(* IEC 61131-3 sources: SortJet_MasterSPS_Aufbau.fbsproj/Device.device.xml.v3^/Plc Logic.plclogic.xml.v3^/Application.application.xml.v3^/09_Station/Stationen/Anlegetisch[201,205]/0_Konfig, 6 files *)

(* ---- Antriebsinformationen_201.gvl ---- *)
(* METADATA
{
	"v3Meta": {
		"objectGuid": "6db4b2f7-21ef-4267-9852-06546c6f86b1"
	}
}
*)
{attribute 'allow_unqualified_access'}
NAMESPACE Antriebsinformationen_201
VAR_GLOBAL

//-------------------------------------------------------------------------------------------------
// ANTRIEBSINFORMATION
//-------------------------------------------------------------------------------------------------

  apgInfoStation201Glastransport : ARRAY[cWAND_1..cANZAHL_WAENDE] OF AntriebsInformationen := [
    (
      wAchsID                                 :=     13,  // Achs ID aus dem EConSet
      stTyp                                   := 'Belt',  // Typ
      wpSchaltschrank                         :=   2010,  // Daten aus dem Schaltplan
      wpSchaltplanreihe                       :=      2,  // Daten aus dem Schaltplan
      wpSchaltplanseite                       :=    100,  // Daten aus dem Schaltplan
      rpMaxGeschwindigkeit                    :=   1000,  // [mm/s]   Max- Geschwindigkeit für den Automatikbetrieb
      rpHandGeschwindigkeit                   :=    200,  // [mm/s]   Hand- Geschwindigkeit
      rpReduzierteGeschwindigkeit             :=     67,  // [mm/s]   Reduzierte Geschwindigkeit
      rpReferenzGeschwindigkeit               :=      0,  // [mm/s]   Geschwindigkeit für die Referenzfahrt
      rpEinrichtGeschwindigkeit               :=     50,  // [mm/s]   Max Geschwindigkeit während der Einrichtung der Anlage
      rpMaxBeschleunigung                     :=   1500,  // [mm/s^2] Max Beschleunigung
      rpMaxVerzoegerung                       :=   2000,  // [mm/s^2] Max Verzoegerung
      rpMaxRuckzeit                           :=     50,  // [ms]     Ruckzeit des Antriebs
      rpReduzierteBeschleunigung              :=   1000,  // [mm/s^2] Reduzierte Beschleunigung
      rpReduzierteVerzoegerung                :=   1000,  // [mm/s^2] Reduzierte Verzoegerung
      rpBeschleunigungFremdanlage             :=   1000,  // [mm/s^2] Beschleunigung zu einer Fremdanlage
      rpGeschwindigkeitMessen                 :=    667,  // [mm/s] Geschwindigkeit beim Scheiben messen
      rpGeschwindigkeitSystemcheck            :=  500.0,  // [mm/s]   Geschwindigkeit im Systemcheck (nur Glastransport)
      rpGeschwindigkeitSystemcheckReduzierung :=  167.0,  // [mm/s]   Geschwindigkeit im Systemcheck bei belegtem Vorstop-Sensor (nur Glastransport)
      stOptionen                              := ( eEndschalterQuelle    := Endschalterquelle_EN.KEINE,     // Hardware-Endschalter: KEINE, UMRICHTER oder SPS
                                                   bVersorgungUeberXVR   := FALSE,                          // XVR-Modus: brueckt Hauptschalter 400 V und LS 230 V
                                                   bBremseLoesenFreigabe := FALSE )                         // Der Antrieb darf über eine Betriebsart die Bremse lösen
    )];

  apgInfoStation201Glastransport_Slave : ARRAY[cWAND_1..cANZAHL_WAENDE] OF AntriebsInformationen := [
    (
      wAchsID                                 :=     65,  // Achs ID aus dem EConSet
      stTyp                                   := 'BeltSl',  // Typ
      wpSchaltschrank                         :=      0,  // Daten aus dem Schaltplan
      wpSchaltplanreihe                       :=      2,  // Daten aus dem Schaltplan
      wpSchaltplanseite                       :=    100,  // Daten aus dem Schaltplan
      rpMaxGeschwindigkeit                    :=   1000,  // [mm/s]   Max- Geschwindigkeit für den Automatikbetrieb
      rpHandGeschwindigkeit                   :=    333,  // [mm/s]   Hand- Geschwindigkeit
      rpReduzierteGeschwindigkeit             :=    250,  // [mm/s]   Reduzierte Geschwindigkeit
      rpReferenzGeschwindigkeit               :=      0,  // [mm/s]   Geschwindigkeit für die Referenzfahrt
      rpEinrichtGeschwindigkeit               :=    100,  // [mm/s]   Max Geschwindigkeit während der Einrichtung der Anlage
      rpMaxBeschleunigung                     :=   1500,  // [mm/s^2] Max Beschleunigung
      rpMaxVerzoegerung                       :=   2000,  // [mm/s^2] Max Verzoegerung
      rpMaxRuckzeit                           :=     50,  // [ms]     Ruckzeit des Antriebs
      rpReduzierteBeschleunigung              :=    500,  // [mm/s^2] Reduzierte Beschleunigung
      rpReduzierteVerzoegerung                :=    500,  // [mm/s^2] Reduzierte Verzoegerung
      rpBeschleunigungFremdanlage             :=      0,  // [mm/s^2] Beschleunigung zu einer Fremdanlage
      rpGeschwindigkeitMessen                 :=   1000,  // [mm/s] Geschwindigkeit beim Scheiben messen
      rpGeschwindigkeitSystemcheck            :=  500.0,  // [mm/s]   Geschwindigkeit im Systemcheck (nur Glastransport)
      rpGeschwindigkeitSystemcheckReduzierung :=  167.0,  // [mm/s]   Geschwindigkeit im Systemcheck bei belegtem Vorstop-Sensor (nur Glastransport)
      stOptionen                              := ( eEndschalterQuelle    := Endschalterquelle_EN.KEINE,     // Hardware-Endschalter: KEINE, UMRICHTER oder SPS
                                                   bVersorgungUeberXVR   := FALSE,                          // XVR-Modus: brueckt Hauptschalter 400 V und LS 230 V
                                                   bBremseLoesenFreigabe := FALSE )                         // Der Antrieb darf über eine Betriebsart die Bremse lösen
    )];

  apgInfoStation201Messachse : AntriebsInformationen :=
    (
      wAchsID                                 :=        14,  // Achs ID aus dem EConSet
      stTyp                                   := 'Measure',  // Typ
      wpSchaltschrank                         :=      2011,  // Daten aus dem Schaltplan
      wpSchaltplanreihe                       :=         2,  // Daten aus dem Schaltplan
      wpSchaltplanseite                       :=       100,  // Daten aus dem Schaltplan
      rpMaxGeschwindigkeit                    :=      1000,  // [mm/s]   Max- Geschwindigkeit für den Automatikbetrieb
      rpHandGeschwindigkeit                   :=       333,  // [mm/s]   Hand- Geschwindigkeit
      rpReduzierteGeschwindigkeit             :=         0,  // [mm/s]   Reduzierte Geschwindigkeit
      rpReferenzGeschwindigkeit               :=        50,  // [mm/s]   Geschwindigkeit für die Referenzfahrt
      rpEinrichtGeschwindigkeit               :=         0,  // [mm/s]   Max Geschwindigkeit während der Einrichtung der Anlage
      rpMaxBeschleunigung                     :=      2500,  // [mm/s^2] Max Beschleunigung
      rpMaxVerzoegerung                       :=      2500,  // [mm/s^2] Max Verzoegerung
      rpMaxRuckzeit                           :=       500,  // [ms]     Ruckzeit des Antriebs
      rpReduzierteBeschleunigung              :=       500,  // [mm/s^2] Reduzierte Beschleunigung
      rpReduzierteVerzoegerung                :=       500,  // [mm/s^2] Reduzierte Verzoegerung
      rpBeschleunigungFremdanlage             :=         0,  // [mm/s^2] Beschleunigung zu einer Fremdanlage
      rpGeschwindigkeitMessen                 :=         0,  // [mm/s] Geschwindigkeit beim Scheiben messen
      rpGeschwindigkeitSystemcheck            :=     500.0,  // [mm/s]   Geschwindigkeit im Systemcheck (nur Glastransport)
      rpGeschwindigkeitSystemcheckReduzierung :=     167.0,  // [mm/s]   Geschwindigkeit im Systemcheck bei belegtem Vorstop-Sensor (nur Glastransport)
      stOptionen                              := ( eEndschalterQuelle    := Endschalterquelle_EN.UMRICHTER, // Hardware-Endschalter: KEINE, UMRICHTER oder SPS
                                                   bVersorgungUeberXVR   := FALSE,                          // XVR-Modus: brueckt Hauptschalter 400 V und LS 230 V
                                                   bBremseLoesenFreigabe := FALSE )                         // Der Antrieb darf über eine Betriebsart die Bremse lösen
    );

END_VAR

END_NAMESPACE

(* ---- Antriebsinformationen_205.gvl ---- *)
(* METADATA
{
	"v3Meta": {
		"objectGuid": "115b641a-a462-4b18-943b-f0d19b116a3d"
	}
}
*)
{attribute 'allow_unqualified_access'}
NAMESPACE Antriebsinformationen_205
VAR_GLOBAL

//-------------------------------------------------------------------------------------------------
// ANTRIEBSINFORMATION
//-------------------------------------------------------------------------------------------------

  apgInfoStation205Glastransport : ARRAY[cWAND_1..cANZAHL_WAENDE] OF AntriebsInformationen := [
    (
      wAchsID                                 :=     9,  // Achs ID aus dem EConSet
      stTyp                                   := 'Belt',  // Typ
      wpSchaltschrank                         :=   2050,  // Daten aus dem Schaltplan
      wpSchaltplanreihe                       :=      2,  // Daten aus dem Schaltplan
      wpSchaltplanseite                       :=    100,  // Daten aus dem Schaltplan
      rpMaxGeschwindigkeit                    :=   1000,  // [mm/s]   Max- Geschwindigkeit für den Automatikbetrieb
      rpHandGeschwindigkeit                   :=    200,  // [mm/s]   Hand- Geschwindigkeit
      rpReduzierteGeschwindigkeit             :=     67,  // [mm/s]   Reduzierte Geschwindigkeit
      rpReferenzGeschwindigkeit               :=      0,  // [mm/s]   Geschwindigkeit für die Referenzfahrt
      rpEinrichtGeschwindigkeit               :=     50,  // [mm/s]   Max Geschwindigkeit während der Einrichtung der Anlage
      rpMaxBeschleunigung                     :=   1500,  // [mm/s^2] Max Beschleunigung
      rpMaxVerzoegerung                       :=   2000,  // [mm/s^2] Max Verzoegerung
      rpMaxRuckzeit                           :=     50,  // [ms]     Ruckzeit des Antriebs
      rpReduzierteBeschleunigung              :=   1000,  // [mm/s^2] Reduzierte Beschleunigung
      rpReduzierteVerzoegerung                :=   1000,  // [mm/s^2] Reduzierte Verzoegerung
      rpBeschleunigungFremdanlage             :=   1000,  // [mm/s^2] Beschleunigung zu einer Fremdanlage
      rpGeschwindigkeitMessen                 :=    667,  // [mm/s] Geschwindigkeit beim Scheiben messen
      rpGeschwindigkeitSystemcheck            :=  500.0,  // [mm/s]   Geschwindigkeit im Systemcheck (nur Glastransport)
      rpGeschwindigkeitSystemcheckReduzierung :=  167.0,  // [mm/s]   Geschwindigkeit im Systemcheck bei belegtem Vorstop-Sensor (nur Glastransport)
      stOptionen                              := ( eEndschalterQuelle    := Endschalterquelle_EN.KEINE,     // Hardware-Endschalter: KEINE, UMRICHTER oder SPS
                                                   bVersorgungUeberXVR   := FALSE,                          // XVR-Modus: brueckt Hauptschalter 400 V und LS 230 V
                                                   bBremseLoesenFreigabe := FALSE )                         // Der Antrieb darf über eine Betriebsart die Bremse lösen
    )];

  apgInfoStation205Glastransport_Slave : ARRAY[cWAND_1..cANZAHL_WAENDE] OF AntriebsInformationen := [
    (
      wAchsID                                 :=     65,  // Achs ID aus dem EConSet
      stTyp                                   := 'BeltSl',  // Typ
      wpSchaltschrank                         :=      0,  // Daten aus dem Schaltplan
      wpSchaltplanreihe                       :=      2,  // Daten aus dem Schaltplan
      wpSchaltplanseite                       :=    100,  // Daten aus dem Schaltplan
      rpMaxGeschwindigkeit                    :=   1000,  // [mm/s]   Max- Geschwindigkeit für den Automatikbetrieb
      rpHandGeschwindigkeit                   :=    333,  // [mm/s]   Hand- Geschwindigkeit
      rpReduzierteGeschwindigkeit             :=    250,  // [mm/s]   Reduzierte Geschwindigkeit
      rpReferenzGeschwindigkeit               :=      0,  // [mm/s]   Geschwindigkeit für die Referenzfahrt
      rpEinrichtGeschwindigkeit               :=    100,  // [mm/s]   Max Geschwindigkeit während der Einrichtung der Anlage
      rpMaxBeschleunigung                     :=   1500,  // [mm/s^2] Max Beschleunigung
      rpMaxVerzoegerung                       :=   2000,  // [mm/s^2] Max Verzoegerung
      rpMaxRuckzeit                           :=     50,  // [ms]     Ruckzeit des Antriebs
      rpReduzierteBeschleunigung              :=    500,  // [mm/s^2] Reduzierte Beschleunigung
      rpReduzierteVerzoegerung                :=    500,  // [mm/s^2] Reduzierte Verzoegerung
      rpBeschleunigungFremdanlage             :=      0,  // [mm/s^2] Beschleunigung zu einer Fremdanlage
      rpGeschwindigkeitMessen                 :=   1000,  // [mm/s] Geschwindigkeit beim Scheiben messen
      rpGeschwindigkeitSystemcheck            :=  500.0,  // [mm/s]   Geschwindigkeit im Systemcheck (nur Glastransport)
      rpGeschwindigkeitSystemcheckReduzierung :=  167.0,  // [mm/s]   Geschwindigkeit im Systemcheck bei belegtem Vorstop-Sensor (nur Glastransport)
      stOptionen                              := ( eEndschalterQuelle    := Endschalterquelle_EN.KEINE,     // Hardware-Endschalter: KEINE, UMRICHTER oder SPS
                                                   bVersorgungUeberXVR   := FALSE,                          // XVR-Modus: brueckt Hauptschalter 400 V und LS 230 V
                                                   bBremseLoesenFreigabe := FALSE )                         // Der Antrieb darf über eine Betriebsart die Bremse lösen
    )];

  apgInfoStation205Messachse : AntriebsInformationen :=
    (
      wAchsID                                 :=        10,  // Achs ID aus dem EConSet
      stTyp                                   := 'Measure',  // Typ
      wpSchaltschrank                         :=      2051,  // Daten aus dem Schaltplan
      wpSchaltplanreihe                       :=         2,  // Daten aus dem Schaltplan
      wpSchaltplanseite                       :=       100,  // Daten aus dem Schaltplan
      rpMaxGeschwindigkeit                    :=      1000,  // [mm/s]   Max- Geschwindigkeit für den Automatikbetrieb
      rpHandGeschwindigkeit                   :=       333,  // [mm/s]   Hand- Geschwindigkeit
      rpReduzierteGeschwindigkeit             :=         0,  // [mm/s]   Reduzierte Geschwindigkeit
      rpReferenzGeschwindigkeit               :=        50,  // [mm/s]   Geschwindigkeit für die Referenzfahrt
      rpEinrichtGeschwindigkeit               :=         0,  // [mm/s]   Max Geschwindigkeit während der Einrichtung der Anlage
      rpMaxBeschleunigung                     :=      2500,  // [mm/s^2] Max Beschleunigung
      rpMaxVerzoegerung                       :=      2500,  // [mm/s^2] Max Verzoegerung
      rpMaxRuckzeit                           :=       500,  // [ms]     Ruckzeit des Antriebs
      rpReduzierteBeschleunigung              :=       500,  // [mm/s^2] Reduzierte Beschleunigung
      rpReduzierteVerzoegerung                :=       500,  // [mm/s^2] Reduzierte Verzoegerung
      rpBeschleunigungFremdanlage             :=         0,  // [mm/s^2] Beschleunigung zu einer Fremdanlage
      rpGeschwindigkeitMessen                 :=         0,  // [mm/s] Geschwindigkeit beim Scheiben messen
      rpGeschwindigkeitSystemcheck            :=     500.0,  // [mm/s]   Geschwindigkeit im Systemcheck (nur Glastransport)
      rpGeschwindigkeitSystemcheckReduzierung :=     167.0,  // [mm/s]   Geschwindigkeit im Systemcheck bei belegtem Vorstop-Sensor (nur Glastransport)
      stOptionen                              := ( eEndschalterQuelle    := Endschalterquelle_EN.UMRICHTER, // Hardware-Endschalter: KEINE, UMRICHTER oder SPS
                                                   bVersorgungUeberXVR   := FALSE,                          // XVR-Modus: brueckt Hauptschalter 400 V und LS 230 V
                                                   bBremseLoesenFreigabe := FALSE )                         // Der Antrieb darf über eine Betriebsart die Bremse lösen
    );

END_VAR

END_NAMESPACE

(* ---- MK_Station_201.gvl ---- *)
(* METADATA
{
	"v3Meta": {
		"objectGuid": "3c311fcf-86c3-480c-8d89-6d8c270ee569"
	}
}
*)
{attribute 'allow_unqualified_access'}
NAMESPACE MK_Station_201
VAR_GLOBAL

//-------------------------------------------------------------------------------------------------
// MASCHINEPARAMETER: ANLEGETISCH
//-------------------------------------------------------------------------------------------------

  apgMKStation201 : Parameter_Station :=
    (
      stStationsNummern                     := ( NummerIntern :=   201,                                                      // Stationsnummer fuer das MMI und die Stationsangabe der Meldungen
                                                 NummerExtern :=  1201,                                                      // Stationsnummer fuer Bedienermeldungen
                                                 NummerSPS    :=   201 ),                                                    // Stationsnummer SPS-intern (Indizes)
      bDeaktivieren                         := FALSE,                                                                        // Station deaktiviert (keine Auftraege, keine Referenzfahrt)
      wMeldungsNummer                       := 1700,                                                                         // Basis-Meldungsnummer (WatchIO)
      eStationsTyp                          := eStation,                                                                     // Typ der Station
      eaAutomatikkreis                      := [eAutomatikkreis_1],                                                          // Automatikkreise, zu denen die Station gehoert
      eaSicherheitskreis                    := [eSicherheitskreis_2],                                                        // Sicherheitskreise, in die die Station eingebunden ist
      // astSicherheitskreisTeilabschaltung
      eSystemcheckZyklus                    := eSystemcheckZyklus_1,                                                         // In welchem Zyklus des Systemchecks die Station geprueft wird
      stSchnittstellendaten                 := ( wVorgaengerStation := cSTATION_DEFAULT,                                     // Station vor dieser Station (cSTATION_DYNAMISCH bei mehreren)
                                                 wNachfolgerStation := cSTATION_202,                                         // Station nach dieser Station (cSTATION_DYNAMISCH bei mehreren)
                                                 bStationIstShuttle := FALSE                                                 // Station ist ein Shuttle
                                               ),
      stStationsOptionen                    := ( stSystemcheck   :=  ( bScheibenVermessenSystemCheck               := TRUE,  // Scheiben im Systemcheck vermessen
                                                                       bScheibeNachSystemcheckAufAuslauf           := FALSE, // Scheibe nach dem Systemcheck auf den Auslaufsensor fahren
                                                                       bSystemCheckMitVorgaengerBatchTransport     := FALSE, // derzeit ohne Funktion
                                                                       bSystemCheckMitNachfolgerBatchTransport     := FALSE, // derzeit ohne Funktion
                                                                       bOptionSystemCheckScheibeMittigLegen        := FALSE  // derzeit ohne Funktion
                                                                     ),
                                                 stAnlegetisch   :=  (
                                                                       bIstAnlegestation                         := TRUE,    // Station an der Scheiben angelegt werden [Anlegetisch, Anlegewand]; im Systemcheck-Verbund nur mit genau einer Scheibe
                                                                       bAnschlagAutomatischAusfahren             := TRUE,    // Anschlaege beim Anlegen automatisch ausfahren (Vorgabe, am Taster umschaltbar)
                                                                       bAnlegetischMitEintransportVorgaenger     := FALSE    // VSG: Station entscheidet selbst zwischen Eintransport vom Vorgaenger und Anlegen
                                                                     ),
                                                 // stTransfershuttle
                                                 stGlastransport :=  ( bVortransport                             := FALSE,   // Vortransport aktivieren [Bsp.: Nach einem Eintransport mit gesetztem Bit <Letzte Scheibe>]
                                                                       bTransportMasterSlaveEintransport         := FALSE,   // derzeit ohne Funktion
                                                                       bTransportMasterSlaveAustransport         := TRUE,    // Austransport als Slave auf die Achse des Nachfolgers
                                                                       bGLasUebernahmeSenkrecht                  := FALSE,   // RKT - Eintransport in Senkrechter-Position bzw. in Waagerechter- Position [default]
                                                                       bAustransportISOLinie                     := FALSE,   // Austransport an eine ISO-Linie
                                                                       bScheibenVermessen                        := TRUE,    // Scheibenmessung am Anlegetisch/Anlegewand
                                                                       bMessrichtungNegativ                      := FALSE,   // Negative Fahrtrichtung beim Messen
                                                                       bScheibenmessungEintransport              := FALSE,   // Scheibenmessung beim Eintransport
                                                                       bScheibenmessungSensorVorabAuslauf        := FALSE    // Scheibenmessung mit SensorVorabAuslauf z.B. Anlegewand
                                                                      ),
                                                 // stEckuebergabe
                                                 // stDrehstation
                                                 bVorAbKomponentenAnsteuerung              := FALSE,                         // VorAbKomponentenAnsteuerung Auftraege werden bearbeitet
                                                 bVerstellungEinAusGefahrenLogikDrehen     := FALSE,                         // Verstellung: Logik ein-/ausgefahren gedreht
                                                 bLangsamfahrtNockenQuerfahrtAktivieren    := FALSE,                         // Querfahrt: Langsamfahrt-Nocken auswerten
                                                 bSKBlockierenDurchVorabSensoren           := FALSE,                         // Vorab-Sensoren belegt blockieren das Oeffnen des Sicherheitskreises
                                                 bStationLeerfahrenBeiSkAnforderung        := FALSE,                         // Station bei Anforderung Sicherheitskreis leerfahren
                                                 bGlasAbgenommenAutomatischQuittieren      := FALSE,                         // derzeit ohne Funktion
                                                 bScheibeAbnehmenNachEintransport          := FALSE                          // Scheibe nach dem Eintransport wieder abnehmen
                                               ),
      stStationsAufbau                      := ( bGeblase                      := [ cANZAHL_WAENDE(TRUE) ],                  // Ausbaustufe: Geblaese je Wand
                                                 bGlastransport                := [ cANZAHL_WAENDE(TRUE) ],                  // Ausbaustufe: Glastransport je Wand
                                                 bKippen                       := [ cANZAHL_WAENDE(TRUE) ],                  // Ausbaustufe: Kippen je Wand (Kipptisch 201 laut E-Plan)
                                                 bKippenSchuetz                := FALSE,                                     // Kippen ueber Schuetz statt Umrichter
                                                 bTransportVerstellung         := [ cANZAHL_WAENDE(FALSE) ],                 // Ausbaustufe Shuttle: Transport-/Dickenverstellung je Wand
                                                 bHub                          := FALSE,                                     // Ausbaustufe: Hub der Station
                                                 bHubrahmen                    := TRUE,                                      // Ausbaustufe: Hubrahmen (Riemen heben/senken)
                                                 bDrehen                       := FALSE,                                     // Ausbaustufe: Drehen
                                                 bQuerachse                    := FALSE,                                     // Ausbaustufe: Querachse
                                                 bMessachse                    := TRUE,                                      // Ausbaustufe: Messachse (Anlegetisch, Anlegewand)
                                                 bDruckluft                    := TRUE,                                      // Druckluftueberwachung vorhanden
                                                 bAnschlag                     := TRUE,                                      // Ausbaustufe: Ausrichtanschlaege
                                                 bSensorAuslauf                := TRUE,                                      // Auslaufsensor vorhanden
                                                 bSensorEinlauf                := TRUE,                                      // Einlaufsensor vorhanden
                                                 bSensorEinlaufStopp           := FALSE,                                     // Shuttle: zusaetzlicher Stopp-Sensor am Einlauf (ohne: Einlaufsensor), Gegenstueck zum Auslauf-Stopp im Rueckwaertstransport
                                                 bSensorAuslaufStopp           := FALSE,                                     // Shuttle: zusaetzlicher Stopp-Sensor am Auslauf (ohne: Auslaufsensor), Verfahrfreigabe und Scheibe hat Shuttle verlassen
                                                 bDurchlaufSperreZumNachfolger := FALSE,                                     // Ausbaustufe: bewegliche Abschrankung zum Nachfolger
                                                 bQuerfahrt                    := FALSE,                                     // Ausbaustufe: Querfahrt
                                                 bKipparme                     := FALSE,                                     // Ausbaustufe: Kipparme
                                                 bSlaveAntrieb                 := FALSE,                                     // Glastransport mit Slave-Antrieb
                                                 bMessachseAmEndeVomTisch      := FALSE,                                     // Messachse am Ende des Tisches (Hoehenfehler fragt den Bediener)
                                                 bWandverstellung              := [ FALSE ],                                 // Ausbaustufe Station: Wandverstellung je Wand
                                                 bWandverstellungMotorisch     := FALSE,                                     // Shuttle: Transport-/Wandverstellung mit Antrieb statt pneumatisch
                                                 bRoellchenleiste              := [ FALSE ],                                 // Ausbaustufe Station: Roellchenleiste je Wand
                                                 bDurchgang                    := FALSE,                                     // Station ist Teil eines Durchgangs (belegt = Oeffnen blockiert)
                                                 bRolltor                      := FALSE,                                     // Ausbaustufe Faecherwagen: Rolltor
                                                 bKlemmzylinder                := FALSE,                                     // Ausbaustufe Faecherwagen: Klemmzylinder fixiert den Oberrahmen beim Ein- und Ausschleusen
                                                 bGreifer                      := [cANZAHL_WAENDE(FALSE)],                   // Shuttle: Greifer je Wand (Scheibe aus dem Faecherwagen ziehen bzw. hineinschieben)
                                                 bRFID                         := FALSE,                                     // RFID-Leser vorhanden
                                                 bAGV                          := FALSE,                                     // Ausbaustufe Faecherwagen: Betrieb mit AGV
                                                 bDLSSchmiersystem             := FALSE,                                     // Zentralschmierung DLS vorhanden
                                                 bGlastransportSlaveVorhanden  := FALSE,                                     // Glastransport mit Slave-Antrieb (Meldungen/Ueberwachung Slave)
                                                 wHydraulikstation             := 0                                          // Faecherwagen Hydraulik: zugeordnete Hydraulikstation (cHYDRAULIKSTATION_x), 0 = keine
                                               ),
      stStationsParameter                   := ( rLaengeUebergroesseScheibe              := 4240,                            // Shuttle: ab dieser Scheibenlaenge gilt die Scheibe als uebergross [mm]
                                                 rMinGlasHoeheAutomatischenEintransport  := 500,                             // VSG: Mindesthoehe fuer automatischen Eintransport [mm]
                                                 rMinGlasLaengeAutomatischenEintransport := 500,                             // VSG: Mindestlaenge fuer automatischen Eintransport [mm]
                                                 wMaximaleAnzahlAktiverAuftraege         := 1,                               // derzeit ohne Funktion
                                                 rMinPosSwEsEingrenzung                  := 0.0,                             // Externer zusaetzlicher Software-Endschalter MIN; 0 = inaktiv; darf den MK-MIN nur weiter eingrenzen
                                                 rMaxPosSwEsEingrenzung                  := 0.0,                             // Externer zusaetzlicher Software-Endschalter MAX; 0 = inaktiv; darf den MK-MAX nur weiter eingrenzen
                                                 rPosFreigabePufferAusfahren             := 0.0                              // derzeit ohne Funktion
                                              ),
      // stFremdanlage
      stGlasdaten                           := [(
                                                 rlMinGlasLaenge                  := 350,                                    // minimal zulässige GlasLänge
                                                 rlMaxGlasLaenge                  := 2500,                                   // maximale zulässige GlasLänge
                                                 rlMinGlasHoehe                   := 190,                                    // minimal zulässige GlasHöhe
                                                 rlMaxGlasHoehe                   := 1800,                                   // maximale zulässige GlasHöhe
                                                 rlMinGlasDicke                   := 3,                                    // minimal zulässige GlasDicke
                                                 rlMaxGlasDicke                   := 12.76,                                     // maximal zulaessige Glasdicke [mm]
                                                 rlLaengeMaxGlas                  := 0.0                                     // maximal zulaessige Glaslaenge [mm]
                                               )]
      // astShuttleAnhaltenQuellen
    );

  apgMKStation201Glastransport : ARRAY[cWAND_1..cANZAHL_WAENDE] OF Parameter_Glastransport := [
    (
      rLaengeStation                        := 3200, // Länge der Station
      rScheibenabstand                      :=  300, // Der Abstand zwischen zwei Scheiben auf der Station
      rWegUeberEinlauf                      :=   50, // Weg ueber den Einlaufsensor hinaus [mm]
      rWegUeberAuslauf                      :=   50, // Weg ueber den Auslaufsensor hinaus [mm]
      rWegUeberSensorenSystemCheck          :=   15, // Der Weg der Ueber ein die Sensoren zum vermessen der Scheiben
      rUeberwachungAuslaufsensor            :=  500, // Ueberwachung des Auslaufsensors [Strecke in der der Auslaufsensor Frei / ueberfahren werden soll]
      rUeberwachungEinlaufsensor            :=  500, // Ueberwachung des Einlaufsensors [Strecke in der der Einlaufsensor Frei / ueberfahren werden soll]
      rWegUeberEinlaufEintransport          :=  150, // Eintransport vorwaerts: Abstand Scheibenhinterkante zum Einlaufsensor [mm]
      rWegUeberEinlaufAustransport          :=   50, // Lage Auf Einlauf: Scheibe liegt um diesen Weg auf dem Einlaufsensor [mm]
      rWegUeberAuslaufEintransport          :=   50, // Eintransport rueckwaerts: Abstand Scheibenhinterkante zum Auslaufsensor [mm]
      rWegUeberAuslaufAustransport          :=   50, // Lage Auf Auslauf: Weg ueber den Auslaufsensor hinaus [mm]
      rWegEinlaufsensorZuVorStopSensor      := 3100, // Beschreibt den Weg vum eine Scheibe beim EIntransport vom Einlaufsensor bis ueberden Vorabstopsensor zu verfahren
      rMesstoleranz                         :=   10, // Toleranz-Mass fuer die Scheibenlaengenmessung
      rMessstrecke                          := 3140, // Beschreibt die Strecke ziwischen 2 Sensoren die der Antrieb verfaehrt
      rWegstreckeBisZurVerzoegerung         := 2600  // Beschreibt die Strecke die gefahren werden soll bis der Antrieb abgebremst werden soll, dies gilt fuer Eintransportauftraege die das Bit "Letzte Scheibe" gesetzt haben
    )];

  apgMKStation201Messachse : Parameter_Messachse :=
    (
      rPositionUeberScheibenhoehe           :=      0, // Position der Zentrierleiste ueber dem Glas so dass das Glas angelegt werden kann
      rKorrekturOffset                      :=      0, // Korrektur der Position um einen Bestimmten Wert (Offset)
      rStreckePositionieren                 :=      0, // ?
      rVerfahrbereichsOffset                :=      0, // Korrektur des Verfahrens wenn
      rOffsetMessung                        :=      0, // ?
      rToleranz                             :=     10, // Toleranzwert in der Ausmessung der Höhe
      rAbstandSensorenOberUndUnterkante     :=    153, // Rechnerischer Abstand zwischen dem Sensor der die Scheibenunterkante misst und dem Sensor der die Scheibenoberkante misst
      rKorrekturOffsetVSGEintransport       := 0.0,    // Korrektur der Position um einen Bestimmten Wert (Offset) beim Eintransport von VSG
      rOffsetNullLinie                      := 0.0     // Offset das auf den Wert des Abstands zur Null-Linie aufgerechnet wird, um dies evtl zu korrigieren
    );

END_VAR
END_NAMESPACE

(* ---- MK_Station_205.gvl ---- *)
(* METADATA
{
	"v3Meta": {
		"objectGuid": "7b970d81-93e6-42b4-b0eb-c486128876da"
	}
}
*)
{attribute 'allow_unqualified_access'}
NAMESPACE MK_Station_205
VAR_GLOBAL

//-------------------------------------------------------------------------------------------------
// MASCHINEPARAMETER: ANLEGETISCH
//-------------------------------------------------------------------------------------------------

  apgMKStation205 : Parameter_Station :=
    (
      stStationsNummern                     := ( NummerIntern :=   205,                                                      // Stationsnummer fuer das MMI und die Stationsangabe der Meldungen
                                                 NummerExtern :=  1205,                                                      // Stationsnummer fuer Bedienermeldungen
                                                 NummerSPS    :=   205 ),                                                    // Stationsnummer SPS-intern (Indizes)
      bDeaktivieren                         := FALSE,                                                                         // Station deaktiviert (keine Auftraege, keine Referenzfahrt)
      wMeldungsNummer                       := 1760,                                                                         // Basis-Meldungsnummer (WatchIO)
      eStationsTyp                          := eStation,                                                                     // Typ der Station
      eaAutomatikkreis                      := [eAutomatikkreis_1],                                                          // Automatikkreise, zu denen die Station gehoert
      eaSicherheitskreis                    := [eSicherheitskreis_Undefiniert],                                              // Sicherheitskreise, in die die Station eingebunden ist
      // astSicherheitskreisTeilabschaltung
      eSystemcheckZyklus                    := eSystemcheckZyklus_1,                                                         // In welchem Zyklus des Systemchecks die Station geprueft wird
      stSchnittstellendaten                 := ( wVorgaengerStation := cSTATION_501,                                         // Station vor dieser Station (cSTATION_DYNAMISCH bei mehreren)
                                                 wNachfolgerStation := cSTATION_204,                                         // Station nach dieser Station (cSTATION_DYNAMISCH bei mehreren)
                                                 bStationIstShuttle := FALSE                                                 // Station ist ein Shuttle
                                               ),
      stStationsOptionen                    := ( stSystemcheck   :=  ( bScheibenVermessenSystemCheck               := TRUE,  // Scheiben im Systemcheck vermessen
                                                                       bScheibeNachSystemcheckAufAuslauf           := FALSE, // Scheibe nach dem Systemcheck auf den Auslaufsensor fahren
                                                                       bSystemCheckMitVorgaengerBatchTransport     := FALSE, // derzeit ohne Funktion
                                                                       bSystemCheckMitNachfolgerBatchTransport     := FALSE, // derzeit ohne Funktion
                                                                       bOptionSystemCheckScheibeMittigLegen        := FALSE  // derzeit ohne Funktion
                                                                     ),
                                                 stAnlegetisch   :=  (
                                                                       bIstAnlegestation                         := TRUE,    // Station an der Scheiben angelegt werden [Anlegetisch, Anlegewand]; im Systemcheck-Verbund nur mit genau einer Scheibe
                                                                       bAnschlagAutomatischAusfahren             := TRUE,    // Anschlaege beim Anlegen automatisch ausfahren (Vorgabe, am Taster umschaltbar)
                                                                       bAnlegetischMitEintransportVorgaenger     := TRUE     // VSG: Station entscheidet selbst zwischen Eintransport vom Vorgaenger und Anlegen
                                                                     ),
                                                 // stTransfershuttle
                                                 stGlastransport :=  ( bVortransport                             := FALSE,   // Vortransport aktivieren [Bsp.: Nach einem Eintransport mit gesetztem Bit <Letzte Scheibe>]
                                                                       bTransportMasterSlaveEintransport         := FALSE,   // derzeit ohne Funktion
                                                                       bTransportMasterSlaveAustransport         := TRUE,    // Austransport als Slave auf die Achse des Nachfolgers
                                                                       bGLasUebernahmeSenkrecht                  := FALSE,   // RKT - Eintransport in Senkrechter-Position bzw. in Waagerechter- Position [default]
                                                                       bAustransportISOLinie                     := FALSE,   // Austransport an eine ISO-Linie
                                                                       bScheibenVermessen                        := TRUE,    // Scheibenmessung am Anlegetisch/Anlegewand
                                                                       bMessrichtungNegativ                      := FALSE,   // Negative Fahrtrichtung beim Messen
                                                                       bScheibenmessungEintransport              := FALSE,   // Scheibenmessung beim Eintransport
                                                                       bScheibenmessungSensorVorabAuslauf        := FALSE    // Scheibenmessung mit SensorVorabAuslauf z.B. Anlegewand
                                                                      ),
                                                 // stEckuebergabe
                                                 // stDrehstation
                                                 bVorAbKomponentenAnsteuerung              := FALSE,                         // VorAbKomponentenAnsteuerung Auftraege werden bearbeitet
                                                 bVerstellungEinAusGefahrenLogikDrehen     := FALSE,                         // Verstellung: Logik ein-/ausgefahren gedreht
                                                 bLangsamfahrtNockenQuerfahrtAktivieren    := FALSE,                         // Querfahrt: Langsamfahrt-Nocken auswerten
                                                 bSKBlockierenDurchVorabSensoren           := FALSE,                         // Vorab-Sensoren belegt blockieren das Oeffnen des Sicherheitskreises
                                                 bStationLeerfahrenBeiSkAnforderung        := FALSE,                         // Station bei Anforderung Sicherheitskreis leerfahren
                                                 bGlasAbgenommenAutomatischQuittieren      := FALSE,                         // derzeit ohne Funktion
                                                 bScheibeAbnehmenNachEintransport          := FALSE                          // Scheibe nach dem Eintransport wieder abnehmen
                                               ),
      stStationsAufbau                      := ( bGeblase                      := [ cANZAHL_WAENDE(TRUE) ],                  // Ausbaustufe: Geblaese je Wand
                                                 bGlastransport                := [ cANZAHL_WAENDE(TRUE) ],                  // Ausbaustufe: Glastransport je Wand
                                                 bKippen                       := [ cANZAHL_WAENDE(FALSE) ],                 // Ausbaustufe: Kippen je Wand (kein Kipptisch an 205)
                                                 bKippenSchuetz                := FALSE,                                     // Kippen ueber Schuetz statt Umrichter
                                                 bTransportVerstellung         := [ cANZAHL_WAENDE(FALSE) ],                 // Ausbaustufe Shuttle: Transport-/Dickenverstellung je Wand
                                                 bHub                          := FALSE,                                     // Ausbaustufe: Hub der Station
                                                 bHubrahmen                    := TRUE,                                      // Ausbaustufe: Hubrahmen (Riemen heben/senken)
                                                 bDrehen                       := FALSE,                                     // Ausbaustufe: Drehen
                                                 bQuerachse                    := FALSE,                                     // Ausbaustufe: Querachse
                                                 bMessachse                    := TRUE,                                      // Ausbaustufe: Messachse (Anlegetisch, Anlegewand)
                                                 bDruckluft                    := TRUE,                                      // Druckluftueberwachung vorhanden
                                                 bAnschlag                     := TRUE,                                      // Ausbaustufe: Ausrichtanschlaege
                                                 bSensorAuslauf                := TRUE,                                      // Auslaufsensor vorhanden
                                                 bSensorEinlauf                := TRUE,                                      // Einlaufsensor vorhanden
                                                 bSensorEinlaufStopp           := FALSE,                                     // Shuttle: zusaetzlicher Stopp-Sensor am Einlauf (ohne: Einlaufsensor), Gegenstueck zum Auslauf-Stopp im Rueckwaertstransport
                                                 bSensorAuslaufStopp           := FALSE,                                     // Shuttle: zusaetzlicher Stopp-Sensor am Auslauf (ohne: Auslaufsensor), Verfahrfreigabe und Scheibe hat Shuttle verlassen
                                                 bDurchlaufSperreZumNachfolger := FALSE,                                     // Ausbaustufe: bewegliche Abschrankung zum Nachfolger
                                                 bQuerfahrt                    := FALSE,                                     // Ausbaustufe: Querfahrt
                                                 bKipparme                     := FALSE,                                     // Ausbaustufe: Kipparme
                                                 bSlaveAntrieb                 := FALSE,                                     // Glastransport mit Slave-Antrieb
                                                 bMessachseAmEndeVomTisch      := FALSE,                                     // Messachse am Ende des Tisches (Hoehenfehler fragt den Bediener)
                                                 bWandverstellung              := [ FALSE ],                                 // Ausbaustufe Station: Wandverstellung je Wand
                                                 bWandverstellungMotorisch     := FALSE,                                     // Shuttle: Transport-/Wandverstellung mit Antrieb statt pneumatisch
                                                 bRoellchenleiste              := [ FALSE ],                                 // Ausbaustufe Station: Roellchenleiste je Wand
                                                 bDurchgang                    := FALSE,                                     // Station ist Teil eines Durchgangs (belegt = Oeffnen blockiert)
                                                 bRolltor                      := FALSE,                                     // Ausbaustufe Faecherwagen: Rolltor
                                                 bKlemmzylinder                := FALSE,                                     // Ausbaustufe Faecherwagen: Klemmzylinder fixiert den Oberrahmen beim Ein- und Ausschleusen
                                                 bGreifer                      := [cANZAHL_WAENDE(FALSE)],                   // Shuttle: Greifer je Wand (Scheibe aus dem Faecherwagen ziehen bzw. hineinschieben)
                                                 bRFID                         := FALSE,                                     // RFID-Leser vorhanden
                                                 bAGV                          := FALSE,                                     // Ausbaustufe Faecherwagen: Betrieb mit AGV
                                                 bDLSSchmiersystem             := FALSE,                                     // Zentralschmierung DLS vorhanden
                                                 bGlastransportSlaveVorhanden  := FALSE,                                     // Glastransport mit Slave-Antrieb (Meldungen/Ueberwachung Slave)
                                                 wHydraulikstation             := 0                                          // Faecherwagen Hydraulik: zugeordnete Hydraulikstation (cHYDRAULIKSTATION_x), 0 = keine
                                               ),
      stStationsParameter                   := ( rLaengeUebergroesseScheibe              := 4240,                            // Shuttle: ab dieser Scheibenlaenge gilt die Scheibe als uebergross [mm]
                                                 rMinGlasHoeheAutomatischenEintransport  := 500,                             // VSG: Mindesthoehe fuer automatischen Eintransport [mm]
                                                 rMinGlasLaengeAutomatischenEintransport := 500,                             // VSG: Mindestlaenge fuer automatischen Eintransport [mm]
                                                 wMaximaleAnzahlAktiverAuftraege         := 1,                               // derzeit ohne Funktion
                                                 rMinPosSwEsEingrenzung                  := 0.0,                             // Externer zusaetzlicher Software-Endschalter MIN; 0 = inaktiv; darf den MK-MIN nur weiter eingrenzen
                                                 rMaxPosSwEsEingrenzung                  := 0.0,                             // Externer zusaetzlicher Software-Endschalter MAX; 0 = inaktiv; darf den MK-MAX nur weiter eingrenzen
                                                 rPosFreigabePufferAusfahren             := 0.0                              // derzeit ohne Funktion
                                              ),
      // stFremdanlage
      stGlasdaten                           := [(
                                                 rlMinGlasLaenge                  := 190,                                    // minimal zulässige GlasLänge
                                                 rlMaxGlasLaenge                  := 1800,                                   // maximale zulässige GlasLänge
                                                 rlMinGlasHoehe                   := 350,                                    // minimal zulässige GlasHöhe
                                                 rlMaxGlasHoehe                   := 2500,                                   // maximale zulässige GlasHöhe
                                                 rlMinGlasDicke                   := 3,                                    // minimal zulässige GlasDicke
                                                 rlMaxGlasDicke                   := 12.76,                                     // maximal zulaessige Glasdicke [mm]
                                                 rlLaengeMaxGlas                  := 0.0                                     // maximal zulaessige Glaslaenge [mm]
                                               )]
      // astShuttleAnhaltenQuellen
    );

  apgMKStation205Glastransport : ARRAY[cWAND_1..cANZAHL_WAENDE] OF Parameter_Glastransport := [
    (
      rLaengeStation                        := 2000, // Länge der Station
      rScheibenabstand                      :=  300, // Der Abstand zwischen zwei Scheiben auf der Station
      rWegUeberEinlauf                      :=   50, // Weg ueber den Einlaufsensor hinaus [mm]
      rWegUeberAuslauf                      :=   50, // Weg ueber den Auslaufsensor hinaus [mm]
      rWegUeberSensorenSystemCheck          :=   15, // Der Weg der Ueber ein die Sensoren zum vermessen der Scheiben
      rUeberwachungAuslaufsensor            :=  500, // Ueberwachung des Auslaufsensors [Strecke in der der Auslaufsensor Frei / ueberfahren werden soll]
      rUeberwachungEinlaufsensor            :=  500, // Ueberwachung des Einlaufsensors [Strecke in der der Einlaufsensor Frei / ueberfahren werden soll]
      rWegUeberEinlaufEintransport          :=  150, // Eintransport vorwaerts: Abstand Scheibenhinterkante zum Einlaufsensor [mm]
      rWegUeberEinlaufAustransport          :=   50, // Lage Auf Einlauf: Scheibe liegt um diesen Weg auf dem Einlaufsensor [mm]
      rWegUeberAuslaufEintransport          :=   50, // Eintransport rueckwaerts: Abstand Scheibenhinterkante zum Auslaufsensor [mm]
      rWegUeberAuslaufAustransport          :=   50, // Lage Auf Auslauf: Weg ueber den Auslaufsensor hinaus [mm]
      rWegEinlaufsensorZuVorStopSensor      := 1750, // Beschreibt den Weg vum eine Scheibe beim EIntransport vom Einlaufsensor bis ueberden Vorabstopsensor zu verfahren
      rMesstoleranz                         :=   10, // Toleranz-Mass fuer die Scheibenlaengenmessung
      rMessstrecke                          := 1800, // Beschreibt die Strecke ziwischen 2 Sensoren die der Antrieb verfaehrt
      rWegstreckeBisZurVerzoegerung         := 1200  // Beschreibt die Strecke die gefahren werden soll bis der Antrieb abgebremst werden soll, dies gilt fuer Eintransportauftraege die das Bit "Letzte Scheibe" gesetzt haben
    )];

  apgMKStation205Messachse : Parameter_Messachse :=
    (
      rPositionUeberScheibenhoehe           :=      0, // Position der Zentrierleiste ueber dem Glas so dass das Glas angelegt werden kann
      rKorrekturOffset                      :=      0, // Korrektur der Position um einen Bestimmten Wert (Offset)
      rStreckePositionieren                 :=      0, // ?
      rVerfahrbereichsOffset                :=      0, // Korrektur des Verfahrens wenn
      rOffsetMessung                        :=      0, // ?
      rToleranz                             :=     10, // Toleranzwert in der Ausmessung der Höhe
      rAbstandSensorenOberUndUnterkante     :=    153, // Rechnerischer Abstand zwischen dem Sensor der die Scheibenunterkante misst und dem Sensor der die Scheibenoberkante misst
      rKorrekturOffsetVSGEintransport       := 0.0,    // Korrektur der Position um einen Bestimmten Wert (Offset) beim Eintransport von VSG
      rOffsetNullLinie                      := 0.0     // Offset das auf den Wert des Abstands zur Null-Linie aufgerechnet wird, um dies evtl zu korrigieren
    );

END_VAR
END_NAMESPACE

(* ---- Konfiguration_201.gvl ---- *)
(* METADATA
{
	"v3Meta": {
		"objectGuid": "96545533-c4ac-453b-9299-b2ad8d3a4e76"
	}
}
*)
{attribute 'allow_unqualified_access'}
NAMESPACE Konfiguration_201
VAR_CONFIG

  // Taster
  Globale_Bausteine.Anlegetisch201.in_bKnebelRiemenVor                                   AT %IX6.1    : BOOL; // IO-L - 201 Riemen vor
  Globale_Bausteine.Anlegetisch201.in_bKnebelRiemenZurueck                               AT %IX6.2    : BOOL; // IO-L - 201 Riemen zurueck
  Globale_Bausteine.Anlegetisch201.in_bTasterQuittierungScheibenmessung                  AT %IX6.0    : BOOL; // IO-L - 201 quittieren Fehlmessung
  Globale_Bausteine.Anlegetisch201.in_bTasterGlasAngelegt                                AT %IX6.4  : BOOL; // IO-L - 201 Austransport Start
  Globale_Bausteine.Anlegetisch201.in_bTasterGlasBruch                                   AT %IX6.3    : BOOL; // IO-L - 201 Glasbruch
  Globale_Bausteine.Anlegetisch201.in_bTasterGlasAbgenommen                              AT %MX1.0    : BOOL; // OPTION
  Globale_Bausteine.Anlegetisch201.in_bTasterAnschlaege                                  AT %MX1.0    : BOOL; // OPTION - Taster Anschlaege

  Globale_Bausteine.Anlegetisch201.out_bSignalTasterScheibeAnlegen                       AT %QX6.0    : BOOL; // IO-L - 201 Austransport Start Meldung
  Globale_Bausteine.Anlegetisch201.out_bSignalTasterScheibeQuittieren                    AT %QX5.6    : BOOL; // IO-L - 201 Fehlmessung Scheibe ausgeloest
  Globale_Bausteine.Anlegetisch201.out_bSignalScheibeGlasbruch                           AT %QX5.7    : BOOL; // IO-L - 201 Glasbruch Meldung (wird nicht beschrieben)
  Globale_Bausteine.Anlegetisch201.out_bAmpelSignalRot                                   AT %QX5.5    : BOOL; // IO-L - 201 Stoerung im Betriebsablauf Ampel rot
  Globale_Bausteine.Anlegetisch201.out_bAmpelSignalGruenScheibeAnlegen                   AT %QX5.3    : BOOL; // IO-L - 201 Freigabe Scheibe anlegen Ampel gruen
  Globale_Bausteine.Anlegetisch201.out_bAmpelSignalGlastransportAktiv                    AT %MX2010.2 : BOOL; // OPTION - Ampel Glastransport aktiv
  //Glasbruch QX3.0

  // Gebläse
  Globale_Bausteine.Anlegetisch201.in_bMotorschutzGeblaese_Ok                            AT %IX1.1    : BOOL; // IO-L - 201 Geblaese Sanftstarter / Sicherung OK
  Globale_Bausteine.Anlegetisch201.in_bDrehzahlErreicht                                  AT %IX1.4    : BOOL; // IO-L - 201 Geblaese BY-PASSED
  Globale_Bausteine.Anlegetisch201.in_bTasterGeblaese1Ein                                AT %IX4.7    : BOOL; // IO-L - 201 Taster Geblaese ein
  Globale_Bausteine.Anlegetisch201.in_bTasterGeblaese2Ein                                AT %MX1.0    : BOOL; // OPTION

  Globale_Bausteine.Anlegetisch201.out_bGeblaese1Ein                                     AT %QX0.6    : BOOL; // IO-L - 201 Geblaese einschalten
  Globale_Bausteine.Anlegetisch201.out_bGeblaese2Ein                                     AT %MX2010.3 : BOOL; // OPTION

  // Kippen//SKquittieren_OP IX4.4
  // Kippen//SKquittieren_LTR IX6.0
  Globale_Bausteine.Anlegetisch201.in_bTasterAnforderungKippen                           AT %IX6.5    : BOOL; // IO-L - 201 Anforderung Durchgang nicht Bedienseite
  Globale_Bausteine.Anlegetisch201.in_bTasterAnforderungKippen_OP                        AT %IX3.2    : BOOL; // IO-L - 201 Anforderung Durchgang (OP1)
  Globale_Bausteine.Anlegetisch201.in_bTasterKippenAuf                                   AT %IX6.6    : BOOL; // IO-L - 201 auf nicht Bedienseite
  Globale_Bausteine.Anlegetisch201.in_bTasterKippenAb                                    AT %IX6.7    : BOOL; // IO-L - 201 ab nicht Bedienseite
  Globale_Bausteine.Anlegetisch201.in_bTasterKippenAuf_OP                                AT %IX3.3    : BOOL; // IO-L - 201 auf (OP1)
  Globale_Bausteine.Anlegetisch201.in_bTasterKippenAb_OP                                 AT %IX3.4    : BOOL; // IO-L - 201 ab (OP1)
  Globale_Bausteine.Anlegetisch201.in_bSensorKipptischOben                               AT %IX4.6    : BOOL; // IO-L - 201 Kipptisch oben
  Globale_Bausteine.Anlegetisch201.in_bSensorKippsicherungGeschlossen                    AT %IX4.5    : BOOL; // IO-L - 201 Kippsicherung geschlossen
  Globale_Bausteine.Anlegetisch201.in_bSensorKippsicherungOffen                          AT %IX4.4    : BOOL; // IO-L - 201 Kippsicherung offen
  Globale_Bausteine.Anlegetisch201.in_bSchaltleisteAusgeloest                            AT %IX10.7   : BOOL; // IO-L - 201 Schaltleiste ausgeloest
  Globale_Bausteine.Anlegetisch201.in_bMotorschutzHydraulik                              AT %IX1.6    : BOOL; // IO-L - 201 Hydraulik Motorstarter / Sicherung OK

  //Kippen angefordert_OP  QX1.6
  //Kippen angefordert_LTR QX2.0
  Globale_Bausteine.Anlegetisch201.out_bKipptischAuf                                     AT %QX10.0   : BOOL; // IO-L - 201 kippen auf
  Globale_Bausteine.Anlegetisch201.out_bKipptischAb                                      AT %QX10.1   : BOOL; // IO-L - 201 kippen ab
  Globale_Bausteine.Anlegetisch201.out_bKippsicherungoeffnen                             AT %QX10.2   : BOOL; // IO-L - 201 Kippsicherung oeffnen
  Globale_Bausteine.Anlegetisch201.out_bLeuchteKipptischOffen                            AT %QX6.1    : BOOL; // IO-L - 201 nicht geschlossen nicht Bedienseite
  Globale_Bausteine.Anlegetisch201.out_bLeuchteKipptischOffen_OP                         AT %QX3.2    : BOOL; // IO-L - 201 nicht geschlossen (OP1)
  Globale_Bausteine.Anlegetisch201.out_bHydraulikpumpeEin                                AT %QX1.0    : BOOL; // IO-L - 201 Start Motor Hydraulikpumpe
  Globale_Bausteine.Anlegetisch201.out_bHydraulikpumpeUmlaufVentil                       AT %MX2011.2 : BOOL; // OPTION
  Globale_Bausteine.Anlegetisch201.out_bSchaltleisteAusgeloest                           AT %MX2011.3 : BOOL; // OPTION
  Globale_Bausteine.Anlegetisch201.out_bKipptischHornWarnsignal                          AT %QX5.2    : BOOL; // IO-L - 201 Kipptisch auf / ab Akustisch
  Globale_Bausteine.Anlegetisch201.out_bKipptischAmpelWarnsignal                         AT %QX5.4    : BOOL; // IO-L - 201 Kipptisch auf / ab Ampel gelb

  // Kipparme
  Globale_Bausteine.Anlegetisch201.in_bMotorschutschalterKipparme                        AT %MX1.1    : BOOL; // OPTION
  Globale_Bausteine.Anlegetisch201.in_bTasterKipparmeAuf                                 AT %MX1.0    : BOOL; // OPTION
  Globale_Bausteine.Anlegetisch201.in_bTasterKipparmeAb                                  AT %MX1.0    : BOOL; // OPTION
  Globale_Bausteine.Anlegetisch201.in_bSensorKipparmeAnschlaegeUnten                     AT %MX1.0    : BOOL; // OPTION
  Globale_Bausteine.Anlegetisch201.in_bSensorKipparmeAnschlaegeOben                      AT %MX1.0    : BOOL; // OPTION
  Globale_Bausteine.Anlegetisch201.in_bSensorKipparmeNichtOben                           AT %MX1.0    : BOOL; // OPTION
  Globale_Bausteine.Anlegetisch201.in_bSensorKipparmeNichtUnten                          AT %MX1.0    : BOOL; // OPTION

  Globale_Bausteine.Anlegetisch201.out_bKipparmeAuf                                      AT %MX2011.6 : BOOL; // OPTION
  Globale_Bausteine.Anlegetisch201.out_bKipparmeAb                                       AT %MX2011.7 : BOOL; // OPTION
  Globale_Bausteine.Anlegetisch201.out_bKipparmeAnschlaegeAuf                            AT %MX2012.0 : BOOL; // OPTION
  Globale_Bausteine.Anlegetisch201.out_bKipparmeAnschlaegeAb                             AT %MX2012.1 : BOOL; // OPTION

  // Geblaese-Baustein (Motorschutz und Ausgang kommen von der Station)
  Globale_Bausteine.Anlegetisch201.Geblaese.in_bMotorschutzschalter_OK                            AT %MX1.1   : BOOL; // OPTION
  Globale_Bausteine.Anlegetisch201.Geblaese.out_bStarteGeblaese                                   AT %MX2012.2 : BOOL; // OPTION

END_VAR

END_NAMESPACE

(* ---- Konfiguration_205.gvl ---- *)
(* METADATA
{
	"v3Meta": {
		"objectGuid": "ce58a66a-e378-4c22-8896-4face4c434b8"
	}
}
*)
{attribute 'allow_unqualified_access'}
NAMESPACE Konfiguration_205
VAR_CONFIG

  // Taster
  Globale_Bausteine.Anlegetisch205.in_bKnebelRiemenVor                                   AT %IX7.4    : BOOL; // IO-L - 205 Riemen vor
  Globale_Bausteine.Anlegetisch205.in_bKnebelRiemenZurueck                               AT %IX7.5    : BOOL; // IO-L - 205 Riemen zurueck
  Globale_Bausteine.Anlegetisch205.in_bTasterQuittierungScheibenmessung                  AT %IX7.3    : BOOL; // IO-L - 205 LTR-K quittieren Fehlmessung
  Globale_Bausteine.Anlegetisch205.in_bTasterGlasAngelegt                                AT %MX1.0    : BOOL; // OPTION - Start Eintransport kommt vom Fusstaster am Umrichter
  Globale_Bausteine.Anlegetisch205.in_bTasterGlasBruch                                   AT %IX7.6    : BOOL; // IO-L - 205 Glasbruch
  Globale_Bausteine.Anlegetisch205.in_bTasterGlasAbgenommen                              AT %MX1.0    : BOOL; // OPTION
  Globale_Bausteine.Anlegetisch205.in_bTasterAnschlaege                                  AT %MX1.0    : BOOL; // OPTION

  Globale_Bausteine.Anlegetisch205.out_bSignalTasterScheibeAnlegen                       AT %MX2050.0 : BOOL; // OPTION - Leuchte im weißen Taster Scheibe anlegen
  Globale_Bausteine.Anlegetisch205.out_bSignalTasterScheibeQuittieren                    AT %QX6.4    : BOOL; // IO-L - 205 Fehlmessung Scheibe ausgeloest
  Globale_Bausteine.Anlegetisch205.out_bSignalScheibeGlasbruch                           AT %QX6.5    : BOOL; // IO-L - 205 Glasbruch Meldung (wird nicht beschrieben)
  Globale_Bausteine.Anlegetisch205.out_bAmpelSignalRot                                   AT %MX2050.1 : BOOL; // OPTION - Ampel rot
  Globale_Bausteine.Anlegetisch205.out_bAmpelSignalGruenScheibeAnlegen                   AT %MX2051.5 : BOOL; // OPTION - Ampel laeuft ueber die Umrichter-IOs
  Globale_Bausteine.Anlegetisch205.out_bAmpelSignalGlastransportAktiv                    AT %MX2050.2 : BOOL; // OPTION - Ampel Glastransport aktiv
  //Glasbruch QX3.0

  // Gebläse
  Globale_Bausteine.Anlegetisch205.in_bMotorschutzGeblaese_Ok                            AT %IX1.2    : BOOL; // IO-L - 205 Geblaese Sanftstarter / Sicherung OK
  Globale_Bausteine.Anlegetisch205.in_bDrehzahlErreicht                                  AT %IX1.5    : BOOL; // IO-L - 205 Geblaese BY-PASSED
  Globale_Bausteine.Anlegetisch205.in_bTasterGeblaese1Ein                                AT %IX7.2    : BOOL; // IO-L - 205 Geblaese ein
  Globale_Bausteine.Anlegetisch205.in_bTasterGeblaese2Ein                                AT %MX1.0    : BOOL; // OPTION

  Globale_Bausteine.Anlegetisch205.out_bGeblaese1Ein                                     AT %QX0.7    : BOOL; // IO-L - 205 Geblaese einschalten
  Globale_Bausteine.Anlegetisch205.out_bGeblaese2Ein                                     AT %MX2050.3 : BOOL; // OPTION

  // Kippen//SKquittieren_OP IX4.4
  // Kippen//SKquittieren_LTR IX6.0
  Globale_Bausteine.Anlegetisch205.in_bTasterAnforderungKippen                           AT %MX1.0    : BOOL; // OPTION
  Globale_Bausteine.Anlegetisch205.in_bTasterAnforderungKippen_OP                        AT %MX1.0    : BOOL; // OPTION
  Globale_Bausteine.Anlegetisch205.in_bTasterKippenAuf                                   AT %MX1.0    : BOOL; // OPTION
  Globale_Bausteine.Anlegetisch205.in_bTasterKippenAb                                    AT %MX1.0    : BOOL; // OPTION
  Globale_Bausteine.Anlegetisch205.in_bTasterKippenAuf_OP                                AT %MX1.0    : BOOL; // OPTION
  Globale_Bausteine.Anlegetisch205.in_bTasterKippenAb_OP                                 AT %MX1.0    : BOOL; // OPTION
  Globale_Bausteine.Anlegetisch205.in_bSensorKipptischOben                               AT %MX1.0    : BOOL; // OPTION
  Globale_Bausteine.Anlegetisch205.in_bSensorKippsicherungGeschlossen                    AT %MX1.1    : BOOL; // OPTION
  Globale_Bausteine.Anlegetisch205.in_bSensorKippsicherungOffen                          AT %MX1.0    : BOOL; // OPTION
  Globale_Bausteine.Anlegetisch205.in_bSchaltleisteAusgeloest                            AT %MX1.0    : BOOL; // OPTION
  Globale_Bausteine.Anlegetisch205.in_bMotorschutzHydraulik                              AT %MX1.1    : BOOL; // OPTION

  //Kippen angefordert_OP  QX1.6
  //Kippen angefordert_LTR QX2.0
  Globale_Bausteine.Anlegetisch205.out_bKipptischAuf                                     AT %MX2051.6 : BOOL; // OPTION
  Globale_Bausteine.Anlegetisch205.out_bKipptischAb                                      AT %MX2051.7 : BOOL; // OPTION
  Globale_Bausteine.Anlegetisch205.out_bKippsicherungoeffnen                             AT %MX2052.0 : BOOL; // OPTION
  Globale_Bausteine.Anlegetisch205.out_bLeuchteKipptischOffen                            AT %MX2052.1 : BOOL; // OPTION
  Globale_Bausteine.Anlegetisch205.out_bLeuchteKipptischOffen_OP                         AT %MX2052.2 : BOOL; // OPTION
  Globale_Bausteine.Anlegetisch205.out_bHydraulikpumpeEin                                AT %MX2052.3 : BOOL; // OPTION
  Globale_Bausteine.Anlegetisch205.out_bHydraulikpumpeUmlaufVentil                       AT %MX2050.4 : BOOL; // OPTION
  Globale_Bausteine.Anlegetisch205.out_bSchaltleisteAusgeloest                           AT %MX2050.5 : BOOL; // OPTION
  Globale_Bausteine.Anlegetisch205.out_bKipptischHornWarnsignal                          AT %MX2050.6 : BOOL; // OPTION
  Globale_Bausteine.Anlegetisch205.out_bKipptischAmpelWarnsignal                         AT %MX2050.7 : BOOL; // OPTION

  // Kipparme
  Globale_Bausteine.Anlegetisch205.in_bMotorschutschalterKipparme                        AT %MX1.1    : BOOL; // OPTION
  Globale_Bausteine.Anlegetisch205.in_bTasterKipparmeAuf                                 AT %MX1.0    : BOOL; // OPTION
  Globale_Bausteine.Anlegetisch205.in_bTasterKipparmeAb                                  AT %MX1.0    : BOOL; // OPTION
  Globale_Bausteine.Anlegetisch205.in_bSensorKipparmeAnschlaegeUnten                     AT %MX1.0    : BOOL; // OPTION
  Globale_Bausteine.Anlegetisch205.in_bSensorKipparmeAnschlaegeOben                      AT %MX1.0    : BOOL; // OPTION
  Globale_Bausteine.Anlegetisch205.in_bSensorKipparmeNichtOben                           AT %MX1.0    : BOOL; // OPTION
  Globale_Bausteine.Anlegetisch205.in_bSensorKipparmeNichtUnten                          AT %MX1.0    : BOOL; // OPTION

  Globale_Bausteine.Anlegetisch205.out_bKipparmeAuf                                      AT %MX2051.0 : BOOL; // OPTION
  Globale_Bausteine.Anlegetisch205.out_bKipparmeAb                                       AT %MX2051.1 : BOOL; // OPTION
  Globale_Bausteine.Anlegetisch205.out_bKipparmeAnschlaegeAuf                            AT %MX2051.2 : BOOL; // OPTION
  Globale_Bausteine.Anlegetisch205.out_bKipparmeAnschlaegeAb                             AT %MX2051.3 : BOOL; // OPTION

  // Geblaese-Baustein (Motorschutz und Ausgang kommen von der Station)
  Globale_Bausteine.Anlegetisch205.Geblaese.in_bMotorschutzschalter_OK                            AT %MX1.1   : BOOL; // OPTION
  Globale_Bausteine.Anlegetisch205.Geblaese.out_bStarteGeblaese                                   AT %MX2051.4 : BOOL; // OPTION

END_VAR

END_NAMESPACE
